Fanuc KAREL source: KB00112.KL

PROGRAM KB00112
%NOLOCKGROUP
VAR
  P1: JOINTPOS
  RESULT: BOOLEAN
BEGIN
  RESULT = J_IN_RANGE(P1)
END KB00112
